(* PLC project MixTank_MT01, Siemens AG TIA Portal V18 Update 3, author j.berger *)
(* stored: creationDateTime 2026-08-27T10:41:12, contentDescription Mixing tank MT01 - FB_Mixer (LAD), FC_ScaleAnalog (SCL), version 1.4, modificationDateTime 2026-08-27T10:41:12, organization Plant 2 - Utilities, language en-US *)
(* Mixing tank MT01, CPU 1214C DC/DC/DC (6ES7214-1AG40-0XB0, firmware V4.6) with SM 1231 AI4 (6ES7231-4HD32-0XB0). *)

(* Scale a 4-20 mA analog input word to engineering units with wire-break detection. *)
FUNCTION FC_ScaleAnalog : REAL
  VAR_INPUT
    Raw : INT;  (* Analog input word (S7 format) *)
    LoEng : REAL;  (* Engineering value at 4 mA *)
    HiEng : REAL;  (* Engineering value at 20 mA *)
  END_VAR
  VAR_OUTPUT
    Fault : BOOL;  (* Wire break or out of range *)
  END_VAR
  VAR_TEMP
    Norm : REAL;  (* Normalised value 0..1 *)
  END_VAR

            // Scale an S7 analog input word from a 4-20 mA channel to engineering units.
// S7-1200 nominal range for 4-20 mA: 4 mA = 0, 20 mA = 27648; overrange up to 32511,
// 32767 (16#7FFF) = wire break / overflow, -4864 = underrange limit.
IF #Raw > 32511 OR #Raw < -4864 THEN
    #Fault := TRUE;
    #FC_ScaleAnalog := #LoEng;
    RETURN;
END_IF;
#Fault := FALSE;

// Normalise raw counts to 0.0 .. 1.0
#Norm := NORM_X(MIN := 0, VALUE := #Raw, MAX := 32767);

// Engineering units
#FC_ScaleAnalog := SCALE_X(MIN := #LoEng, VALUE := #Norm, MAX := #HiEng);

          
END_FUNCTION

(* Mixing tank MT01 batch sequence, interlocks and alarms. *)
FUNCTION_BLOCK FB_Mixer
  VAR
    S_Idle : BOOL := TRUE;  (* Step: idle, ready for start *)
    S_FillA : BOOL;  (* Step: fill ingredient A *)
    S_FillB : BOOL;  (* Step: fill ingredient B *)
    S_Heat : BOOL;  (* Step: heat with agitation *)
    S_Mix : BOOL;  (* Step: timed mix at temperature *)
    S_Drain : BOOL;  (* Step: drain tank *)
    S_Done : BOOL;  (* Step: batch complete, wait for acknowledge *)
    Fault : BOOL;  (* Any alarm active *)
    Alm_EStop : BOOL;  (* Alarm: emergency stop *)
    Alm_AgitOverload : BOOL;  (* Alarm: agitator motor overload *)
    Alm_HeaterOvertemp : BOOL;  (* Alarm: heater safety thermostat tripped *)
    Alm_LevelHH : BOOL;  (* Alarm: tank level high-high *)
    Alm_LevelSensor : BOOL;  (* Alarm: level transmitter wire break / out of range *)
    Alm_TempSensor : BOOL;  (* Alarm: temperature transmitter wire break / out of range *)
    Alm_AgitFeedback : BOOL;  (* Alarm: agitator commanded but no running feedback *)
    Alm_FillTimeout : BOOL;  (* Alarm: filling took longer than 10 min *)
    Level_Pct : REAL;  (* Tank level, % *)
    Temp_C : REAL;  (* Tank temperature, degC *)
    Level_Fault : BOOL;  (* Level input out of range *)
    Temp_Fault : BOOL;  (* Temperature input out of range *)
    Level_Above_Min : BOOL;  (* Level above agitator / heater minimum *)
    SP_Level_A : REAL := 40.0;  (* Setpoint: level after ingredient A, % *)
    SP_Level_B : REAL := 80.0;  (* Setpoint: level after ingredient B, % *)
    SP_Temp : REAL := 65.0;  (* Setpoint: batch temperature, degC *)
    Agit_Min_Level : REAL := 20.0;  (* Minimum level for agitator and heater, % *)
    SP_Drain_Empty : REAL := 3.0;  (* Level considered empty when draining, % *)
    Mix_Time : TIME := T#5M;  (* Mix time at temperature *)
    Batch_Count : INT;  (* Completed batches *)
    T_AgitFB : TON;  (* Agitator feedback watchdog *)
    T_FillTimeout : TON;  (* Fill watchdog *)
    T_Mix : TON;  (* Mix timer *)
    T_DrainDelay : TON;  (* Drain run-on after empty *)
    C_Batch : CTU;  (* Batch counter *)
  END_VAR
  VAR_EXTERNAL
    Start_PB : BOOL;  (* Start pushbutton S1 (NO) *)
    Stop_PB : BOOL;  (* Stop pushbutton S2 (NC, TRUE = not pressed) *)
    EStop_OK : BOOL;  (* E-stop safety relay K0 OK *)
    Agitator_Running : BOOL;  (* Agitator contactor K3 auxiliary contact (running feedback) *)
    Agitator_OL_OK : BOOL;  (* Agitator motor protector Q3 not tripped *)
    LSHH_OK : BOOL;  (* High-high level switch LSHH101 (NC, TRUE = level not high-high) *)
    Outlet_Valve_Closed : BOOL;  (* Outlet valve XV103 closed limit switch *)
    Lid_Closed : BOOL;  (* Tank lid / manway closed switch *)
    Reset_PB : BOOL;  (* Reset / acknowledge pushbutton S3 (NO) *)
    Heater_OT_OK : BOOL;  (* Heater safety thermostat TSH102 OK (not over-temperature) *)
    Inlet_Valve_A : BOOL;  (* Ingredient A (water) inlet valve XV101 *)
    Inlet_Valve_B : BOOL;  (* Ingredient B (syrup) inlet valve XV102 *)
    Outlet_Valve : BOOL;  (* Outlet / drain valve XV103 *)
    Agitator_Run : BOOL;  (* Agitator motor M1 contactor K3 *)
    Heater_On : BOOL;  (* Immersion heater E1 contactor K4 *)
    Lamp_Running : BOOL;  (* Batch running lamp H1 (green) *)
    Lamp_Fault : BOOL;  (* Fault lamp H2 (red) *)
    Lamp_Batch_Done : BOOL;  (* Batch complete lamp H3 (white) *)
    Level_Raw : INT;  (* Level transmitter LT101, 4-20 mA = 0-100 % (SM 1231 ch0, raw 0..27648) *)
    Temp_Raw : INT;  (* Temperature transmitter TT101, 4-20 mA = 0-150 degC (SM 1231 ch1, raw 0..27648) *)
    HMI_Reset_Count : BOOL;  (* HMI button: reset batch counter *)
  END_VAR
  VAR  (* added by the conversion: wires and edge detectors of the diagram *)
    _FC_ScaleAnalog3_Fault : ANY;
    _FC_ScaleAnalog3_OUT : REAL;
    _FC_ScaleAnalog12_Fault : ANY;
    _FC_ScaleAnalog12_OUT : REAL;
    R_TRIG1 : R_TRIG;
    _GE122_ENO : BOOL;
    _GE122_OUT : BOOL;
    _GE131_ENO : BOOL;
    _GE131_OUT : BOOL;
    _GE140_ENO : BOOL;
    _GE140_OUT : BOOL;
    _LE157_ENO : BOOL;
    _LE157_OUT : BOOL;
    _LT214_ENO : BOOL;
    _LT214_OUT : BOOL;
  END_VAR

(* LD diagram, written out as Structured Text *)
(* Scale level transmitter LT101 (4-20 mA -> 0-100 %) *)
_FC_ScaleAnalog3_OUT := FC_ScaleAnalog(Raw := Level_Raw, LoEng := 0.0, HiEng := 100.0, Fault => _FC_ScaleAnalog3_Fault);
Level_Pct := _FC_ScaleAnalog3_OUT;
Level_Fault := _FC_ScaleAnalog3_Fault;
(* Scale temperature transmitter TT101 (4-20 mA -> 0-150 degC) *)
_FC_ScaleAnalog12_OUT := FC_ScaleAnalog(Raw := Temp_Raw, LoEng := 0.0, HiEng := 150.0, Fault => _FC_ScaleAnalog12_Fault);
Temp_C := _FC_ScaleAnalog12_OUT;
Temp_Fault := _FC_ScaleAnalog12_Fault;
(* Level above minimum for agitator and heater *)
Level_Above_Min := Level_Pct >= Agit_Min_Level;
(* Alarm: Emergency stop pressed *)
IF NOT EStop_OK THEN Alm_EStop := TRUE; END_IF;
(* Alarm: Agitator motor overload *)
IF NOT Agitator_OL_OK THEN Alm_AgitOverload := TRUE; END_IF;
(* Alarm: Heater safety thermostat tripped *)
IF NOT Heater_OT_OK THEN Alm_HeaterOvertemp := TRUE; END_IF;
(* Alarm: Tank level high-high *)
IF NOT LSHH_OK THEN Alm_LevelHH := TRUE; END_IF;
(* Alarm: Level transmitter fault *)
IF Level_Fault THEN Alm_LevelSensor := TRUE; END_IF;
(* Alarm: Temperature transmitter fault *)
IF Temp_Fault THEN Alm_TempSensor := TRUE; END_IF;
(* Alarm: Agitator no running feedback *)
T_AgitFB(IN := Agitator_Run AND NOT Agitator_Running, PT := T#3S);
IF T_AgitFB.Q THEN Alm_AgitFeedback := TRUE; END_IF;
(* Alarm: Fill timeout *)
T_FillTimeout(IN := S_FillA OR S_FillB, PT := T#10M);
IF T_FillTimeout.Q THEN Alm_FillTimeout := TRUE; END_IF;
(* Acknowledge alarms (conditions still present set again) *)
IF Reset_PB THEN Alm_EStop := FALSE; END_IF;
IF Reset_PB THEN Alm_AgitOverload := FALSE; END_IF;
IF Reset_PB THEN Alm_HeaterOvertemp := FALSE; END_IF;
IF Reset_PB THEN Alm_LevelHH := FALSE; END_IF;
IF Reset_PB THEN Alm_LevelSensor := FALSE; END_IF;
IF Reset_PB THEN Alm_TempSensor := FALSE; END_IF;
IF Reset_PB THEN Alm_AgitFeedback := FALSE; END_IF;
IF Reset_PB THEN Alm_FillTimeout := FALSE; END_IF;
(* Fault summary *)
Fault := Alm_EStop OR Alm_AgitOverload OR Alm_HeaterOvertemp OR Alm_LevelHH OR Alm_LevelSensor OR Alm_TempSensor OR Alm_AgitFeedback OR Alm_FillTimeout;
(* Stop or fault: abort batch, back to idle *)
IF NOT Stop_PB OR Fault THEN S_FillA := FALSE; END_IF;
IF NOT Stop_PB OR Fault THEN S_FillB := FALSE; END_IF;
IF NOT Stop_PB OR Fault THEN S_Heat := FALSE; END_IF;
IF NOT Stop_PB OR Fault THEN S_Mix := FALSE; END_IF;
IF NOT Stop_PB OR Fault THEN S_Drain := FALSE; END_IF;
IF NOT Stop_PB OR Fault THEN S_Done := FALSE; END_IF;
IF NOT Stop_PB OR Fault THEN S_Idle := TRUE; END_IF;
(* Idle -> Fill A: start with outlet closed and lid closed *)
R_TRIG1(CLK := Start_PB);
IF S_Idle AND R_TRIG1.Q AND Stop_PB AND NOT Fault AND Outlet_Valve_Closed AND Lid_Closed THEN S_Idle := FALSE; END_IF;
IF S_Idle AND R_TRIG1.Q AND Stop_PB AND NOT Fault AND Outlet_Valve_Closed AND Lid_Closed THEN S_FillA := TRUE; END_IF;
(* Fill A -> Fill B at level setpoint A *)
_GE122_OUT := GE(EN := S_FillA, IN1 := Level_Pct, IN2 := SP_Level_A, ENO => _GE122_ENO);
IF _GE122_OUT THEN S_FillA := FALSE; END_IF;
IF _GE122_OUT THEN S_FillB := TRUE; END_IF;
(* Fill B -> Heat at level setpoint B *)
_GE131_OUT := GE(EN := S_FillB, IN1 := Level_Pct, IN2 := SP_Level_B, ENO => _GE131_ENO);
IF _GE131_OUT THEN S_FillB := FALSE; END_IF;
IF _GE131_OUT THEN S_Heat := TRUE; END_IF;
(* Heat -> Mix at temperature setpoint *)
_GE140_OUT := GE(EN := S_Heat, IN1 := Temp_C, IN2 := SP_Temp, ENO => _GE140_ENO);
IF _GE140_OUT THEN S_Heat := FALSE; END_IF;
IF _GE140_OUT THEN S_Mix := TRUE; END_IF;
(* Mix for Mix_Time, then drain *)
T_Mix(IN := S_Mix, PT := Mix_Time);
IF T_Mix.Q THEN S_Mix := FALSE; END_IF;
IF T_Mix.Q THEN S_Drain := TRUE; END_IF;
(* Drain until empty plus 10 s *)
_LE157_OUT := LE(EN := S_Drain, IN1 := Level_Pct, IN2 := SP_Drain_Empty, ENO => _LE157_ENO);
T_DrainDelay(IN := _LE157_OUT, PT := T#10S);
IF T_DrainDelay.Q THEN S_Drain := FALSE; END_IF;
IF T_DrainDelay.Q THEN S_Done := TRUE; END_IF;
(* Count completed batches *)
C_Batch(CU := S_Done, R := HMI_Reset_Count, PV := 9999);
Batch_Count := C_Batch.CV;
(* Done -> Idle on acknowledge *)
IF S_Done AND Reset_PB THEN S_Done := FALSE; END_IF;
IF S_Done AND Reset_PB THEN S_Idle := TRUE; END_IF;
(* Inlet valve A *)
Inlet_Valve_A := S_FillA AND NOT Fault AND LSHH_OK AND Outlet_Valve_Closed;
(* Inlet valve B *)
Inlet_Valve_B := S_FillB AND NOT Fault AND LSHH_OK AND Outlet_Valve_Closed;
(* Agitator: heat and mix steps, overload OK, lid closed, level above minimum *)
Agitator_Run := (S_Heat OR S_Mix) AND NOT Fault AND Agitator_OL_OK AND Lid_Closed AND Level_Above_Min;
(* Heater: heat and mix steps, agitator running, level above minimum, thermostat OK, below setpoint *)
_LT214_OUT := LT(EN := (S_Heat OR S_Mix) AND NOT Fault AND Agitator_Running AND Level_Above_Min AND Heater_OT_OK, IN1 := Temp_C, IN2 := SP_Temp, ENO => _LT214_ENO);
Heater_On := _LT214_OUT;
(* Outlet valve *)
Outlet_Valve := S_Drain AND NOT Fault;
(* Running lamp *)
Lamp_Running := S_FillA OR S_FillB OR S_Heat OR S_Mix OR S_Drain;
(* Fault lamp *)
Lamp_Fault := Fault;
(* Batch done lamp *)
Lamp_Batch_Done := S_Done;
END_FUNCTION_BLOCK

CONFIGURATION PLC_1
  RESOURCE PLC_1 ON PLC
    VAR_GLOBAL  (* Default tag table *)
      Start_PB AT %I0.0 : BOOL;  (* Start pushbutton S1 (NO) *)
      Stop_PB AT %I0.1 : BOOL;  (* Stop pushbutton S2 (NC, TRUE = not pressed) *)
      EStop_OK AT %I0.2 : BOOL;  (* E-stop safety relay K0 OK *)
      Agitator_Running AT %I0.3 : BOOL;  (* Agitator contactor K3 auxiliary contact (running feedback) *)
      Agitator_OL_OK AT %I0.4 : BOOL;  (* Agitator motor protector Q3 not tripped *)
      LSHH_OK AT %I0.5 : BOOL;  (* High-high level switch LSHH101 (NC, TRUE = level not high-high) *)
      Outlet_Valve_Closed AT %I0.6 : BOOL;  (* Outlet valve XV103 closed limit switch *)
      Lid_Closed AT %I0.7 : BOOL;  (* Tank lid / manway closed switch *)
      Reset_PB AT %I1.0 : BOOL;  (* Reset / acknowledge pushbutton S3 (NO) *)
      Heater_OT_OK AT %I1.1 : BOOL;  (* Heater safety thermostat TSH102 OK (not over-temperature) *)
      Inlet_Valve_A AT %Q0.0 : BOOL;  (* Ingredient A (water) inlet valve XV101 *)
      Inlet_Valve_B AT %Q0.1 : BOOL;  (* Ingredient B (syrup) inlet valve XV102 *)
      Outlet_Valve AT %Q0.2 : BOOL;  (* Outlet / drain valve XV103 *)
      Agitator_Run AT %Q0.3 : BOOL;  (* Agitator motor M1 contactor K3 *)
      Heater_On AT %Q0.4 : BOOL;  (* Immersion heater E1 contactor K4 *)
      Lamp_Running AT %Q0.5 : BOOL;  (* Batch running lamp H1 (green) *)
      Lamp_Fault AT %Q0.6 : BOOL;  (* Fault lamp H2 (red) *)
      Lamp_Batch_Done AT %Q0.7 : BOOL;  (* Batch complete lamp H3 (white) *)
      Level_Raw AT %IW96 : INT;  (* Level transmitter LT101, 4-20 mA = 0-100 % (SM 1231 ch0, raw 0..27648) *)
      Temp_Raw AT %IW98 : INT;  (* Temperature transmitter TT101, 4-20 mA = 0-150 degC (SM 1231 ch1, raw 0..27648) *)
      HMI_Reset_Count AT %M10.0 : BOOL;  (* HMI button: reset batch counter *)
    END_VAR
    TASK Main(PRIORITY := 1);
    PROGRAM Mixer_DB WITH Main : FB_Mixer;
  END_RESOURCE
END_CONFIGURATION
